Fanuc KAREL source: kt00307.KL

-- PROVISIONAL review KL for V1013-1; original PC SHA256 b09a7c0bc66a124b2f51f5e132a371ac80982898c54c456f807f9d8023650e91
-- Incomplete behavior may be omitted. Consult companion uncertainty JSON. Do not deploy.
PROGRAM KT00307
%NOLOCKGROUP
VAR
  I2 : INTEGER
  OUT : BOOLEAN
-- UNRESOLVED_DECL H1 type=002017
BEGIN
  -- UNRESOLVED_PC offsets 5-19; opcodes 2E,22,9D,33,B4
  -- UNRESOLVED_PC offsets 24-35; opcodes 2E,23
  -- UNRESOLVED_PC offsets 40-62; opcodes 22,9D,33,B3,21,58,23
  -- UNRESOLVED_PC offsets 67-71; opcodes 7F
END KT00307
